TYPE ST_PolarIIChamber_OutsideRingServiceCtrl :
STRUCT
	Lift : ST_PolarIIChamber_LiftTopDownServiceCtrl;
	Rotate : ST_PolarIIChamber_OutsideRingRotateServiceCtrl;
END_STRUCT
END_TYPE

(* stored: Version 1.1.0.1, ProductVersion 3.1.4026.18
   DUT ST_PolarIIChamber_OutsideRingServiceCtrl: Id {14000000-0000-0000-0000-000000000067} *)
